Fanuc KAREL source: KA00119.KL

PROGRAM KA00119
%NOLOCKGROUP
VAR
  SRC: CONFIG
  DST: ARRAY[2] OF BYTE
BEGIN
  SRC.CFG_FLIP = TRUE
  DST[1] = SRC
END KA00119
